Fanuc KAREL source: KO00016.KL

PROGRAM KO00016
%NOLOCKGROUP
VAR
  P1: XYZWPR
  P2: XYZWPR
  P3: XYZWPR
  P4: XYZWPR
  OUT: JOINTPOS
BEGIN
  OUT = FRAME(P1, P2, P3, P4)
END KO00016
